Staubli VAL3: Lab2B_IsmaL2.dtx


